// TIA Portal V18 export
// export: Created 2026-11-25T00:00:00.0000000Z, ExportSetting WithDefaults
Screen "Setup"  800x480, Number=4
  ScreenLayer 
    TextField "Title" at 8,8 size 600x28  Text="Setup / rig check"
    TextField "LRig" at 8,50 size 420x30  Text="Rig check required (3 rejects in a row)"
    IOField "VRig" at 440,50 size 140x30  FormatPattern=9, Mode=Output
      ProcessValue := RigCheck
    TextField "Step1" at 8,100 size 780x30  Text="1. Put the master part in and run it."
    TextField "Step2" at 8,136 size 780x30  Text="2. Press the acknowledge key at the station. The start stays blocked until then."
